PROGRAM ladder
VAR
	xoutput: BOOL;
	xtest: BOOL;
	xtest2: BOOL;
END_VAR

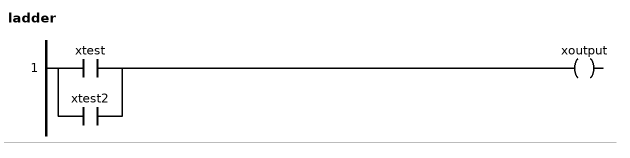
// NETWORK 1
xoutput := xtest OR xtest2;

END_PROGRAM

(* stored: Version 1.1.0.1, ProductVersion 3.1.4024.16
   POU ladder: Id {04d867c5-831f-4a2c-a8ba-57738ccf38e1}, SpecialFunc None *)
